(*
SPDX-License-Identifier: MIT
License: https://opensource.org/license/mit
*)

(*!
<summary>Intentionally omits child-array storage to exercise group validation.</summary>
<description>
Negative fixture: Children intentionally returns an invalid reference without callbacks or exceptions.
Owns no child array or test instances. Use only in the hosting regression task.
</description>
*)

{attribute 'no_assign'}
{attribute 'no_explicit_call' := 'do not call this function block directly'}
FUNCTION_BLOCK MissingChildrenTestGroup EXTENDS TOF_Testing.TestGroup<1>
VAR_STAT
	//! <summary>Class name shared by all instances of this function block.</summary>
	{attribute 'hide'}
	_ClassName : STRING := __POUNAME();
END_VAR
VAR
	{attribute 'hide'}
	{attribute 'init_namespace'}
	_NamespaceName : STRING;
END_VAR

//! <summary>Borrows the concrete class name for the lifetime of this instance; callers must not modify it.</summary>
{attribute 'monitoring' := 'call'}
PROPERTY ClassName : REFERENCE TO STRING
GET
ClassName REF= _ClassName;
END_GET
END_PROPERTY

//! <summary>Borrows the compiler-initialized namespace; callers must not modify the returned reference.</summary>
{attribute 'monitoring' := 'call'}
PROPERTY NamespaceName : REFERENCE TO STRING
GET
NamespaceName REF= _NamespaceName;
END_GET
END_PROPERTY

//! <summary>Reports the complete concrete instance size, excluding separately allocated storage.</summary>
{attribute 'monitoring' := 'call'}
PROPERTY SelfSize : ULINT
GET
SelfSize := XSIZEOF(THIS^);
END_GET
END_PROPERTY

//! <summary>Returns an invalid reference intentionally to exercise missing-storage diagnostics.</summary>
{attribute 'monitoring' := 'call'}
PROPERTY Children : REFERENCE TO ARRAY [0.._ChildCount - 1] OF TOF_Testing.ITestElement
GET
RETURN;
END_GET
END_PROPERTY

END_FUNCTION_BLOCK

(* stored: Version 1.1.0.1
   POU MissingChildrenTestGroup: Id {fb95ab59-a9a2-40ad-938a-0fa0457f6ced}, SpecialFunc None
   Property ClassName: Id {0bd6dd02-ac76-4254-bddc-873df5a9616f}
   Get Get: Id {0f2977db-611b-4ba7-94a0-cbacb8ce5f8d}
   Property NamespaceName: Id {bbd4bc15-2ecd-46f6-b772-55f72789d5dd}
   Get Get: Id {cba722d9-8178-4328-9471-56ff9c24efb4}
   Property SelfSize: Id {b034e448-4e2b-4038-aa06-792637ab354a}
   Get Get: Id {31ca6629-40b5-4821-8a8e-5eb7115fad19}
   Property Children: Id {28be966f-affe-4b7e-a07d-f7bb827477c8}
   Get Get: Id {ff635876-ca89-465b-a3bd-4e69660ed6ca} *)
